(*
SPDX-FileCopyrightText: © 2026 Oleksandr Tiutyk <trofimich@gmail.com>
SPDX-License-Identifier: MIT
License: https://opensource.org/license/mit
*)

(*!
<summary>Provides delayed synthetic acquisition and release for Task stopping tests.</summary>
<description>
The scenario owns this manager and injects it into the task explicitly. Configure inputs before Start.
Operations have no hardware effects. A release exception intentionally leaves the synthetic resource held.
Observations are read-only to the scenario. ResetFixture clears them and the simulated state once the task is inactive.
</description>
*)

FUNCTION_BLOCK TaskStoppingResource EXTENDS TOF_Core.Object IMPLEMENTS TOF_Core.IResourceManager
VAR_INPUT
	//! <summary>Throw before acquisition is scheduled.</summary>
	ThrowOnStartAcquire : BOOL;
	//! <summary>Throw after the last acquisition step has marked the resource acquired.</summary>
	ThrowAfterAcquire : BOOL;
	//! <summary>Throw before release is scheduled, retaining the acquired resource.</summary>
	ThrowOnStartRelease : BOOL;
	//! <summary>Injected exceptions throw again when GetMessage is called.</summary>
	ThrowOnGetMessage : BOOL;
END_VAR
VAR_OUTPUT
	//! <summary>Total acquisition requests across runs.</summary>
	AcquireCalls : UINT;
	//! <summary>Total release requests across runs.</summary>
	ReleaseCalls : UINT;
	//! <summary>Completed steps in the current acquisition.</summary>
	AcquireProgress : UINT;
END_VAR
VAR CONSTANT
	//! <summary>Calls needed for a pending acquisition, allowing cancellation before its response.</summary>
	_AcquireSteps : UINT := 3;
	//! <summary>Calls needed after StartRelease to observe asynchronous completion.</summary>
	_ReleaseSteps : UINT := 2;
END_VAR
VAR_STAT
	//! <summary>Class name shared by all instances of this function block.</summary>
	_ClassName : STRING := __POUNAME();
END_VAR
VAR
	_Acquired : BOOL;
	_Acquiring : BOOL;
	_Releasing : BOOL;
	_ReleaseProgress : UINT;
END_VAR

{attribute 'monitoring' := 'call'}
PROPERTY ClassName : REFERENCE TO STRING
GET
ClassName REF= _ClassName;
END_GET
END_PROPERTY

(*!
<summary>Advances one pending synthetic operation.</summary>
<description>
No pending operation means no action. Acquisition failure may occur after ownership was obtained.
</description>
*)
METHOD Execute
IF _Acquiring THEN
	AcquireProgress := AcquireProgress + 1;

	IF AcquireProgress >= _AcquireSteps THEN
		_Acquiring := FALSE;
		_Acquired := TRUE;

		IF ThrowAfterAcquire THEN
			raiseConfiguredFailure(message := "Acquire failure");
		END_IF
	END_IF
ELSIF _Releasing THEN
	_ReleaseProgress := _ReleaseProgress + 1;

	IF _ReleaseProgress >= _ReleaseSteps THEN
		_Releasing := FALSE;
		_Acquired := FALSE;
	END_IF
END_IF
END_METHOD

(*!
<summary>Drains a late acquisition response without starting a new request.</summary>
<description>
Used by the injected task during OnStopping. A late acquired resource remains available for normal release.
</description>
*)
METHOD INTERNAL FinishPendingAcquire : BOOL
IF _Acquiring THEN
	Execute();
END_IF

FinishPendingAcquire := NOT _Acquiring;
END_METHOD

(*!
<summary>Returns the borrowed manager as a synthetic resource.</summary>
<description>
The caller must not delete it.
</description>
*)
METHOD GetResource : TOF_Core.IObject
GetResource := THIS^;
END_METHOD

(*!
<summary>Borrows the test namespace.</summary>
*)
{attribute 'monitoring' := 'call'}
PROPERTY NamespaceName : REFERENCE TO STRING
GET
NamespaceName REF= CurrentNamespace.Name;
END_GET
END_PROPERTY

(*!
<summary>Raises the configured synthetic exception.</summary>
<description>
Used only by test operations, never by FB lifecycle methods. The throwing formatter exercises diagnostic
fallback.
</description>
<param name="message">Text copied into the injected exception.</param>
*)
METHOD PRIVATE raiseConfiguredFailure
VAR_INPUT
	message : WSTRING(255);
END_VAR
VAR
	failure : TOF_Core.StandardException;
	formattingFailure : ThrowingGetMessageException;
END_VAR
IF ThrowOnGetMessage THEN
	formattingFailure.Throw(
		sourceNamespaceName := NamespaceName,
		sourceClassName := ClassName,
		sourcePOUName := __POUNAME(),
		sourcePosition := __POSITION(),
		message := message
	);
ELSE
	failure.Throw(
		sourceNamespaceName := NamespaceName,
		sourceClassName := ClassName,
		sourcePOUName := __POUNAME(),
		sourcePosition := __POSITION(),
		message := message
	);
END_IF
END_METHOD

(*!
<summary>Reports synthetic resource ownership.</summary>
<description>
Side-effect-free and non-throwing.
</description>
*)
{attribute 'monitoring' := 'call'}
PROPERTY ResourceAcquired : BOOL
GET
ResourceAcquired := _Acquired;
END_GET
END_PROPERTY

(*!
<summary>Reports the concrete fixture size.</summary>
*)
{attribute 'monitoring' := 'call'}
PROPERTY SelfSize : ULINT
GET
SelfSize := XSIZEOF(THIS^);
END_GET
END_PROPERTY

(*!
<summary>Restores idle synthetic state and clears all observations.</summary>
<description>
Call only when the driving task is inactive. Clears synthetic ownership even after an injected release failure.
Leaves fault configuration intact and does not perform physical release.
</description>
*)
METHOD INTERNAL ResetFixture
_Acquired := FALSE;
_Acquiring := FALSE;
_Releasing := FALSE;
_ReleaseProgress := 0;
AcquireProgress := 0;
AcquireCalls := 0;
ReleaseCalls := 0;
END_METHOD

(*!
<summary>Requests one delayed acquisition.</summary>
<description>
An injected early exception leaves no pending operation. An already acquired resource is retained.
</description>
*)
METHOD StartAcquire
AcquireCalls := AcquireCalls + 1;

IF ThrowOnStartAcquire THEN
	raiseConfiguredFailure(message := "Acquire failure");
END_IF

IF NOT _Acquired THEN
	AcquireProgress := 0;
	_Acquiring := TRUE;
END_IF
END_METHOD

(*!
<summary>Requests delayed release or throws the configured terminal failure.</summary>
<description>
The task must issue this once. A thrown request deliberately keeps ResourceAcquired TRUE.
</description>
*)
METHOD StartRelease
ReleaseCalls := ReleaseCalls + 1;

IF ThrowOnStartRelease THEN
	raiseConfiguredFailure(message := "Release failure");
END_IF

_ReleaseProgress := 0;
_Releasing := TRUE;
END_METHOD

END_FUNCTION_BLOCK

(* stored: Version 1.1.0.1, ProductVersion 3.1.4026.21
   POU TaskStoppingResource: Id {bc32d584-5f1f-4adf-b270-32dd155806b0}, SpecialFunc None
   Folder Service methods: Id {cb2e2601-1fab-450c-93e0-25b52d8fa414}
   Property ClassName: Id {77412ac9-0bfe-435e-833d-c765ff25c225}
   Get Get: Id {023f6e75-0fb5-4e94-9b0b-b2d4e91dcdd2}
   Method Execute: Id {4cf9df9e-f4cb-4ad7-be3e-c5c3e9682682}
   Method FinishPendingAcquire: Id {281fbd7a-0e8f-4a9b-bb80-83db7f131abc}
   Method GetResource: Id {817447e8-4f8c-46a5-951d-dfad25609566}
   Property NamespaceName: Id {d3d8c026-dd9e-488f-bca0-4af1f8dab693}
   Get Get: Id {378f92c9-9c4d-41d8-9e89-30980962b838}
   Method raiseConfiguredFailure: Id {7c9ba618-ecbe-46c5-a6fd-5b701df8ef89}
   Property ResourceAcquired: Id {7a735f58-5f9a-4c4b-ada5-70f6d92aec2c}
   Get Get: Id {2cdb29da-1d7a-4031-ae3a-061a41cd9aa6}
   Property SelfSize: Id {5cdf1056-cc1a-45be-b2be-d0580af580dd}
   Get Get: Id {74f9c47a-f463-4b97-b9d8-d5fbd7c93d40}
   Method ResetFixture: Id {1cd6381a-8c17-4988-9f27-607e5a67005e}
   Method StartAcquire: Id {33c5f634-9d63-423e-8608-f38410ecbea8}
   Method StartRelease: Id {5f66b414-8aff-4599-aa8e-cdcda4d1c51a} *)
